# EPICS autosave request: iocs/ad/csimdetector-ioc/db/ADCSimDetector_settings.req
$(P)$(R)TimeStep
$(P)$(R)NumTimePoints
$(P)$(R)AcquireTime

file "NDArrayBase_settings.req", P=$(P), R=$(R)
